FUNCTION_BLOCK PRINT_CHECK
  {SET_ATTRIBUTE(OpcUa, DEVICE.SENSOR)}
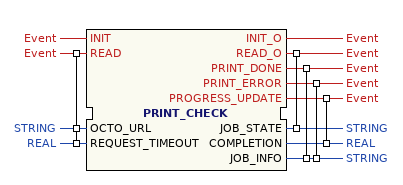
  EVENT_INPUT
    INIT;
    READ WITH OCTO_URL, REQUEST_TIMEOUT;
  END_EVENT
  EVENT_OUTPUT
    INIT_O;
    READ_O WITH JOB_STATE;
    PRINT_DONE WITH JOB_INFO;
    PRINT_ERROR WITH JOB_INFO;
    PROGRESS_UPDATE WITH COMPLETION;
  END_EVENT
  VAR_INPUT
    OCTO_URL : STRING; {SET_ATTRIBUTE(OpcUa, Constant)}
    REQUEST_TIMEOUT : REAL; {SET_ATTRIBUTE(OpcUa, Constant)}
  END_VAR
  VAR_OUTPUT
    JOB_STATE : STRING; {SET_ATTRIBUTE(OpcUa, Variable)}
    COMPLETION : REAL; {SET_ATTRIBUTE(OpcUa, Variable)}
    JOB_INFO : STRING; {SET_ATTRIBUTE(OpcUa, Variable)}
  END_VAR
END_FUNCTION_BLOCK
